Staubli VAL3: _TolleranceCheck.pgx

program _TolleranceCheck(bool& x_bAutoConnect)
  local string l_sMsg
begin

  if bMemState and !isPowered()
    pHere1=here(flange,world)
    l_sMsg="下电位置:"+toString(".2",pHere1.trsf.x)+","+toString(".2",pHere1.trsf.y)+","+toString(".2",pHere1.trsf.rz)
    logMsg(l_sMsg)
    bMemState=false
  elseIf !bMemState and isPowered()
    pHere2=here(flange,world)
    l_sMsg="上电位置:"+toString(".2",pHere1.trsf.x)+","+toString(".2",pHere1.trsf.y)+","+toString(".2",pHere1.trsf.rz)
    logMsg(l_sMsg)
    bMemState=true
  endIf
  //check
  if distance(pHere1.trsf,pHere2.trsf)<10
    x_bAutoConnect=true
  else
    x_bAutoConnect=false
    l_sMsg="TolleranceCheck位置偏差距离过大，需手动连接"
    popUpMsg(l_sMsg)
  endIf

end
